// TIA Portal V20 export
// export: Created 2026-10-19T18:02:57.2651003Z, ExportSetting WithDefaults, DisplayName Totally Integrated Automation Portal, DisplayVersion V20 Update 6, DisplayName TIA Portal Openness, DisplayVersion V20 Update 6, DisplayName TIA Portal Version Control Interface, DisplayVersion V20 Update 6, DisplayName SINAMICS Startdrive Advanced, DisplayVersion V20 SP1, DisplayName SINAMICS Startdrive G130, G150, S120, S150, SINAMICS MV, G220, S200, S210, DisplayVersion V20 SP1, DisplayName SINAMICS Startdrive G110M, G120, G120C, G120D, G120P, G115D, DisplayVersion V20 SP1, DisplayName STEP 7 Professional, DisplayVersion V20 Update 6, DisplayName STEP 7 Safety, DisplayVersion V20 Update 2, DisplayName WinCC Basic/Comfort/Advanced, DisplayVersion V20 Update 6, DisplayName WinCC Unified, DisplayVersion V20 Update 6
DATA_BLOCK "Settings_DB"   // DB71
{ S7_Optimized_Access := 'TRUE' }
VERSION : 0.1
// stored: AutoNumber true, DBAccessibleFromOPCUA true, DBAccessibleFromWebserver true, IsOnlyStoredInLoadMemory false, IsRetainMemResEnabled false, IsWriteProtectedInAS false, MemoryReserve 100
   VAR RETAIN
      Inbound_Cnv_Settings { S7_SetPoint := 'True'} : "Inbound_Cnv_Settings";
      PopUp_Cnv_Settings { S7_SetPoint := 'True'} : Array[1..4] of "PopUp_Cnv_Settings";
      Pick_Cnv_Settings { S7_SetPoint := 'True'} : "Pick_Cnv_Settings";
      Outbound_Cnv_Settings { S7_SetPoint := 'True'} : "Outbound_Cnv_Settings";
      VTD_Settings : "VTD_Settings";
      ECnv_Settings : "ECnv_Settings";
      LCnv_Settings : Array[1..3] of "Buffer_Cnv_Settings";
   END_VAR
   VAR
      "Weighing Station" : Struct
         "Minimum Weight" : Real := 30.0;
         "Maximum Weigh" : Real := 1500.0;
      END_STRUCT;
      "Profile Station" : Struct
         "Maximum Length" : Real := 1230.0;
         "Conveyor Speed mm_s" : Real := 10.0;
      END_STRUCT;
   END_VAR
   VAR RETAIN
      Shuttle_MQTT_Settings : "MQTT_Settings";
      System_Settings : "System_Settings";
   END_VAR
   VAR
      TimeStartBoost_P2ToP3 { S7_SetPoint := 'True'} : UInt := 20;
      TimeStartBoost_P3ToP4 : UInt := 8;
      TimeStartBoost_P1ToP2 : UInt := 8;
   END_VAR
BEGIN
   Inbound_Cnv_Settings.ID := 130001;
   Inbound_Cnv_Settings.TC_Time := 0;
   Inbound_Cnv_Settings.Transfer_Time := 30;
   Inbound_Cnv_Settings.Slow_Speed := 0;
   Inbound_Cnv_Settings.Full_Speed := 60;
   Inbound_Cnv_Settings.Manual_Speed := 60;
   Inbound_Cnv_Settings.No_Forklift_Detect_Timer := 5;
   Inbound_Cnv_Settings.G120_Hardware_ID := 376;
   PopUp_Cnv_Settings[1].ID := 150001;
   PopUp_Cnv_Settings[2].ID := 160001;
   PopUp_Cnv_Settings[3].ID := 170001;
   PopUp_Cnv_Settings[4].ID := 180001;
   PopUp_Cnv_Settings[1..4].Roller_TC_Time := 0;
   PopUp_Cnv_Settings[1..2].Roller_Transfer_Time := 30;
   PopUp_Cnv_Settings[3..4].Roller_Transfer_Time := 25;
   PopUp_Cnv_Settings[1..4].Roller_Slow_Speed := 0;
   PopUp_Cnv_Settings[1..4].Roller_Full_Speed := 60;
   PopUp_Cnv_Settings[1..3].Roller_Manual_Speed := 60;
   PopUp_Cnv_Settings[4].Roller_Manual_Speed := 50;
   PopUp_Cnv_Settings[1..4].Chain_TC_Time := 0;
   PopUp_Cnv_Settings[1].Chain_Transfer_Time := 50;
   PopUp_Cnv_Settings[2].Chain_Transfer_Time := 500;
   PopUp_Cnv_Settings[3].Chain_Transfer_Time := 40;
   PopUp_Cnv_Settings[4].Chain_Transfer_Time := 50;
   PopUp_Cnv_Settings[1..2].Chain_Slow_Speed := 0;
   PopUp_Cnv_Settings[3].Chain_Slow_Speed := 50;
   PopUp_Cnv_Settings[4].Chain_Slow_Speed := 0;
   PopUp_Cnv_Settings[1].Chain_Full_Speed := 60;
   PopUp_Cnv_Settings[2..3].Chain_Full_Speed := 70;
   PopUp_Cnv_Settings[4].Chain_Full_Speed := 60;
   PopUp_Cnv_Settings[1].Chain_Manual_Speed := 30;
   PopUp_Cnv_Settings[2].Chain_Manual_Speed := 60;
   PopUp_Cnv_Settings[3].Chain_Manual_Speed := 50;
   PopUp_Cnv_Settings[4].Chain_Manual_Speed := 60;
   PopUp_Cnv_Settings[1..4].Lift_TC_Time := 0;
   PopUp_Cnv_Settings[1].Lift_Transfer_Time := 7;
   PopUp_Cnv_Settings[2..4].Lift_Transfer_Time := 15;
   PopUp_Cnv_Settings[1..4].Lift_Slow_Speed := 0;
   PopUp_Cnv_Settings[1..2].Lift_Full_Speed := 100;
   PopUp_Cnv_Settings[3].Lift_Full_Speed := 80;
   PopUp_Cnv_Settings[4].Lift_Full_Speed := 100;
   PopUp_Cnv_Settings[1].Lift_Manual_Speed := 40;
   PopUp_Cnv_Settings[2..4].Lift_Manual_Speed := 10;
   PopUp_Cnv_Settings[1].Roller_G120_Hardware_ID := 385;
   PopUp_Cnv_Settings[2].Roller_G120_Hardware_ID := 394;
   PopUp_Cnv_Settings[3].Roller_G120_Hardware_ID := 403;
   PopUp_Cnv_Settings[4].Roller_G120_Hardware_ID := 466;
   PopUp_Cnv_Settings[1].Chain_G120_Hardware_ID := 412;
   PopUp_Cnv_Settings[2].Chain_G120_Hardware_ID := 421;
   PopUp_Cnv_Settings[3].Chain_G120_Hardware_ID := 430;
   PopUp_Cnv_Settings[4].Chain_G120_Hardware_ID := 0;
   PopUp_Cnv_Settings[1].Lift_G120_Hardware_ID := 340;
   PopUp_Cnv_Settings[2].Lift_G120_Hardware_ID := 358;
   PopUp_Cnv_Settings[3].Lift_G120_Hardware_ID := 493;
   PopUp_Cnv_Settings[4].Lift_G120_Hardware_ID := 349;
   Pick_Cnv_Settings.ID := 410001;
   Pick_Cnv_Settings.TC_Time := 0;
   Pick_Cnv_Settings.Transfer_Time := 25;
   Pick_Cnv_Settings.Slow_Speed := 0;
   Pick_Cnv_Settings.Full_Speed := 60;
   Pick_Cnv_Settings.Manual_Speed := 60;
   Pick_Cnv_Settings.No_Forklift_Detect_Timer := 0;
   Pick_Cnv_Settings.G120_Hardware_ID := 412;
   Outbound_Cnv_Settings.ID := 140001;
   Outbound_Cnv_Settings.TC_Time := 0;
   Outbound_Cnv_Settings.Transfer_Time := 25;
   Outbound_Cnv_Settings.Slow_Speed := 0;
   Outbound_Cnv_Settings.Full_Speed := 60;
   Outbound_Cnv_Settings.Manual_Speed := 60;
   Outbound_Cnv_Settings.No_Forklift_Detect_Timer := 5;
   Outbound_Cnv_Settings.G120_Hardware_ID := 367;
   VTD_Settings.ID := 1;
   VTD_Settings.Lowest_Level := 1;
   VTD_Settings.Highest_Level := 3;
   VTD_Settings.VTD_Max_Heigh := 7145;
   VTD_Settings.VTD_Min_Height := 68;
   VTD_Settings.VTD_Level_Granularity := 20;
   VTD_Settings.Dft_Level_Offset_LE := 0;
   VTD_Settings.Dft_Level_Offset_AE := 0;
   VTD_Settings.Teach_Speed := 0;
   VTD_Settings.Creep_Speed := 5;
   VTD_Settings.Slow_Speed := 5;
   VTD_Settings.Slow_Calib_Speed := 5;
   VTD_Settings.Loaded_Speed := 80;
   VTD_Settings.Shuttle_Speed := 80;
   VTD_Settings.Pallet_Speed := 40;
   VTD_Settings.Empty_Speed := 60;
   VTD_Settings.Dock_speed := 5;
   VTD_Settings.Manual_Speed := 10;
   VTD_Settings.Slowdown_Count_LE := 600;
   VTD_Settings.Creep_Count_LE := 60;
   VTD_Settings.Slowdown_Count_AE := 700;
   VTD_Settings.Creep_Count_AE := 60;
   VTD_Settings.Encoder_Delta_W1 := 0.0;
   VTD_Settings.Encoder_Delta_W2 := 0.0;
   VTD_Settings.AE_Ratio := 0.0;
   VTD_Settings.Encoder_Delta_Warning := 60.0;
   VTD_Settings.Encoder_Delta_Error := 80.0;
   VTD_Settings.Transfer_Timeout_Up := 200;
   VTD_Settings.Transfer_Timeout_Down := 200;
   VTD_Settings.Lockpins_Timeout_Extend := 6000;
   VTD_Settings.Lockpins_Timeout_Retract := 6000;
   VTD_Settings.Level_Detect_Timeout := 500;
   VTD_Settings.Teach_Timeout := 600;
   VTD_Settings.Chain_Slack_Timeout := 700;
   VTD_Settings.Level_Detect_LE := 3.0;
   VTD_Settings.G120_Hardware_ID := 612;
   VTD_Settings.Teach_Values.Levels_LE[0] := 69.0;
   VTD_Settings.Teach_Values.Levels_LE[1] := 3451.0;
   VTD_Settings.Teach_Values.Levels_LE[2] := 5249.0;
   VTD_Settings.Teach_Values.Levels_LE[3] := 7049.0;
   VTD_Settings.Teach_Values.Levels_AE[0] := 0;
   VTD_Settings.Teach_Values.Levels_AE[1] := 63;
   VTD_Settings.Teach_Values.Levels_AE[2] := 2069;
   VTD_Settings.Teach_Values.Levels_AE[3] := 4077;
   ECnv_Settings.ID := 120101;
   ECnv_Settings.Barcode_ID := 0;
   ECnv_Settings.Cnv_Level := 1;
   ECnv_Settings.TC_Time := 0;
   ECnv_Settings.Transfer_Time := 20;
   ECnv_Settings.Pallet_Align_Time := 0;
   ECnv_Settings.Slow_Speed := 0;
   ECnv_Settings.Full_Speed := 70;
   ECnv_Settings.Manual_Speed := 50;
   ECnv_Settings.G120_Hardware_ID := 475;
   LCnv_Settings[1].ID := 100101;
   LCnv_Settings[2].ID := 100201;
   LCnv_Settings[3].ID := 100301;
   LCnv_Settings[1..3].Barcode_ID := 0;
   LCnv_Settings[1].Cnv_Level := 1;
   LCnv_Settings[2].Cnv_Level := 2;
   LCnv_Settings[3].Cnv_Level := 3;
   LCnv_Settings[1..3].TC_Time := 1;
   LCnv_Settings[1..3].Transfer_Time := 20;
   LCnv_Settings[1..3].Pallet_Align_Time := 4;
   LCnv_Settings[1..3].Slow_Speed := 25;
   LCnv_Settings[1..3].Full_Speed := 70;
   LCnv_Settings[1..2].Manual_Speed := 60;
   LCnv_Settings[3].Manual_Speed := 50;
   LCnv_Settings[1..3].Safety_stop_Timeout := 0;
   LCnv_Settings[1].G120_Hardware_ID := 439;
   LCnv_Settings[2].G120_Hardware_ID := 448;
   LCnv_Settings[3].G120_Hardware_ID := 457;
   Shuttle_MQTT_Settings.MQTT_Con_Params.hwId := 64;
   Shuttle_MQTT_Settings.MQTT_Con_Params.connId := 16#0001;
   Shuttle_MQTT_Settings.MQTT_Con_Params.broker := '10.0.34.2';
   Shuttle_MQTT_Settings.MQTT_Con_Params.port := 1883;
   Shuttle_MQTT_Settings.MQTT_Con_Params.tls.enableTls := FALSE;
   Shuttle_MQTT_Settings.MQTT_Con_Params.tls.validateServerIdentity := FALSE;
   Shuttle_MQTT_Settings.MQTT_Con_Params.tls.brokerCert := 0;
   Shuttle_MQTT_Settings.MQTT_Con_Params.tls.clientCert := 0;
   Shuttle_MQTT_Settings.MQTT_Con_Params.keepAlive := 60;
   Shuttle_MQTT_Settings.Client_ID := WSTRING#'PLC';
   Shuttle_MQTT_Settings.Username := WSTRING#'Devin';
   Shuttle_MQTT_Settings.Password := WSTRING#'1';
   Shuttle_MQTT_Settings.Timeout := 0;
   Shuttle_MQTT_Settings.QoS := 0;
   Shuttle_MQTT_Settings.Retain := TRUE;
   Shuttle_MQTT_Settings.Will_Topic := WSTRING#'';
   Shuttle_MQTT_Settings.Will_Msg_Length := 0;
   Shuttle_MQTT_Settings.Will_Msg_Payload[1..128] := 16#00;
   System_Settings.VTD_Count := 1;
   System_Settings.Level_Count := 3;
   System_Settings.Cnv_Count := 10;
   System_Settings.Shuttle_Count := 3;
   System_Settings.Shuttle_Interlock_Timeout := 999;
END_DATA_BLOCK
